// TIA Portal project "Impacchettatore" (V18)

(* hardware
DEVICE "S71500/ET200MP station_1"  S7-1500 station
   slot 0: "Telaio di montaggio_0"  Rack  6ES7 590-1***0-0AA0
   slot 1: "PLC_1"  CPU 1516-3 PN/DP  6ES7 516-3AN01-0AB0  V2.5
      slot 3: "Display CPU_1"  6ES7591-1BA00-0AA0
   slot 2: "DI 32x24VDC HF_1"  DI 32x24VDC HF  6ES7 521-1BL00-0AB0  V2.1
   slot 3: "DQ 32x24VDC/0.5A HF_1"  DQ 32x24VDC/0.5A HF  6ES7 522-1BL01-0AB0  V1.0
   slot 4: "AI 8xU/I/RTD/TC ST_1"  AI 8xU/I/RTD/TC ST  6ES7 531-7KF00-0AB0  V2.1
   slot 5: "AQ 4xU/I ST_1"  AQ 4xU/I ST  6ES7 532-5HD00-0AB0  V2.1
*)

// ===== PLC "PLC_1"  CPU 1516-3 PN/DP =====

VAR_GLOBAL   // PLC tag table "Tabella delle variabili standard"
   "slittaCentraleSu" AT %Q0.0 : Bool;
   "slittaCentraleGiu" AT %Q0.1 : Bool;
   "slittaSuperioreAvanti" AT %Q0.2 : Bool;
   "slittaSuperioreIndietro" AT %Q0.3 : Bool;
   "slittaEsternaSu" AT %Q0.4 : Bool;
   "motAvanti" AT %Q0.5 : Bool;
   "hg1" AT %Q0.6 : Bool;
   "hr2" AT %Q0.7 : Bool;
   "sensoreFondo" AT %I0.0 : Bool;
   "sensoreSopra" AT %I0.1 : Bool;
   "marcia" AT %I0.2 : Bool;
   "stop" AT %I0.3 : Bool;
   "inizializzazione" AT %I0.4 : Bool;
   "emergenza" AT %I0.5 : Bool;
   "readSlittaCentraleBasso" AT %I0.6 : Bool;
   "readSlittaCentraleAlto" AT %I0.7 : Bool;
   "readSlittaSuperioreIndietro" AT %I1.0 : Bool;
   "readSlittaSuperioreAvanti" AT %I1.1 : Bool;
   "readSlittaEsternaBasso" AT %I1.2 : Bool;
   "readSlittaEsternaAlto" AT %I1.3 : Bool;
END_VAR

DATA_BLOCK "DB_Comandi"   // DB1
{ S7_Optimized_Access := 'FALSE' }
VERSION : 0.1
   VAR
      btnInizializza : Bool;
      btnResetPezzi : Bool;
      btnStopNastro : Bool;
      btnSlittaLatGiu : Bool;
      btnSlittaLatSu : Bool;
      btnPistoneIndietro : Bool;
      btnPistoneAvanti : Bool;
      btnSlittaCentroGiu : Bool;
      btnSlittaCentroSu : Bool;
      btnNastro : Bool;
      bStop : Bool;
      bAuto : Bool;
      bMan : Bool;
      bReset : Bool;
      bEmergenza : Bool;
   END_VAR
BEGIN
END_DATA_BLOCK

DATA_BLOCK "DB_Stati"   // DB2
{ S7_Optimized_Access := 'FALSE' }
VERSION : 0.1
   VAR
      sAuto : Bool;
      sStop : Bool;
      sMan : Bool;
      sHome : Bool;
      sAttesastop : Bool;
      sEmergenza : Bool;
      bIni1 : Bool;
      bIni2 : Bool;
      bRip1 : Bool;
      bRip2 : Bool;
   END_VAR
BEGIN
END_DATA_BLOCK

DATA_BLOCK "DB_Tappe"   // DB3
{ S7_Optimized_Access := 'FALSE' }
VERSION : 0.1
   VAR
      tappeGemma : Int;
      tappeM1 : Int;
      tappeM2 : Int;
   END_VAR
BEGIN
END_DATA_BLOCK

DATA_BLOCK "DB_Variabili"   // DB4
{ S7_Optimized_Access := 'FALSE' }
VERSION : 0.1
   VAR
      timerResetPulsantiSTART : Bool;
      timerResetPulsantiDONE : Bool;
      timerResetPulsantiOUTPUT : Time;
      timerResetPulsantiDURATA : Time;
      timerSTART_1 : Bool;
      timerDONE_1 : Bool;
      timerOUTPUT_1 : Time;
      timerDURATA_1 : Time;
      timerSTART_2 : Bool;
      timerDONE_2 : Bool;
      timerOUTPUT_2 : Time;
      timerDURATA_2 : Time;
      timerSTART_3 : Bool;
      timerDONE_3 : Bool;
      timerOUTPUT_3 : Time;
      timerDURATA_3 : Time;
      timerSTART_4 : Bool;
      timerDONE_4 : Bool;
      timerOUTPUT_4 : Time;
      timerDURATA_4 : Time;
      statoLED : Bool;
      oSlittaEsterna : Bool;
      oPistoneIndietro : Bool;
      oPistoneAvanti : Bool;
      nCicli : Int;
      nPezzi : Int;
      oNastro : Bool;
      oSlittaSu : Bool;
      oLedVerde : Bool;
      oLedRosso : Bool;
      oSlittaGiu : Bool;
   END_VAR
BEGIN
END_DATA_BLOCK

// folder: System blocks/Program resources

DATA_BLOCK "timerResetPulsanti"   // DB5
{ S7_Optimized_Access := 'TRUE' }
AUTHOR : Simatic
FAMILY : IEC
NAME : IEC_TMR
VERSION : 1.0
// stored: InstanceOfName IEC_TIMER
"IEC_TIMER"
BEGIN
END_DATA_BLOCK

DATA_BLOCK "timer_1"   // DB6
{ S7_Optimized_Access := 'TRUE' }
AUTHOR : Simatic
FAMILY : IEC
NAME : IEC_TMR
VERSION : 1.0
// stored: InstanceOfName IEC_TIMER
"IEC_TIMER"
BEGIN
END_DATA_BLOCK

DATA_BLOCK "timer_2"   // DB7
{ S7_Optimized_Access := 'TRUE' }
AUTHOR : Simatic
FAMILY : IEC
NAME : IEC_TMR
VERSION : 1.0
// stored: InstanceOfName IEC_TIMER
"IEC_TIMER"
BEGIN
END_DATA_BLOCK

DATA_BLOCK "timer_3"   // DB8
{ S7_Optimized_Access := 'TRUE' }
AUTHOR : Simatic
FAMILY : IEC
NAME : IEC_TMR
VERSION : 1.0
// stored: InstanceOfName IEC_TIMER
"IEC_TIMER"
BEGIN
END_DATA_BLOCK

DATA_BLOCK "timer_4"   // DB9
{ S7_Optimized_Access := 'TRUE' }
AUTHOR : Simatic
FAMILY : IEC
NAME : IEC_TMR
VERSION : 1.0
// stored: InstanceOfName IEC_TIMER
"IEC_TIMER"
BEGIN
END_DATA_BLOCK

// folder: (top level)

FUNCTION "FC_Gemma" : Void   // FC1, SCL
{ S7_Optimized_Access := 'TRUE' }
VERSION : 0.1
BEGIN
   CASE "DB_Tappe".tappeGemma OF
       0:  // Stato di stop
           "DB_Stati".sStop := TRUE;
           IF "DB_Comandi".bAuto = TRUE THEN
               "DB_Tappe".tappeGemma := 1; //home
               "DB_Stati".sAttesastop := FALSE;
               "DB_Stati".sAuto := FALSE;
               "DB_Stati".sHome := TRUE;
               "DB_Stati".sMan := FALSE;
               "DB_Stati".sStop := FALSE;
           ELSE
               IF "DB_Comandi".bMan = TRUE THEN
                   "DB_Tappe".tappeGemma := 4; //manuale
                   "DB_Stati".sAttesastop := FALSE;
                   "DB_Stati".sAuto := FALSE;
                   "DB_Stati".sHome := FALSE;
                   "DB_Stati".sMan := TRUE;
                   "DB_Stati".sStop := FALSE;
               END_IF;
           END_IF;
       1:  // Stato di home
           IF "DB_Stati".bIni1 = TRUE AND "DB_Stati".bIni2 = TRUE THEN
               "DB_Tappe".tappeGemma := 2; //automatico
               "DB_Stati".sAttesastop := FALSE;
               "DB_Stati".sAuto := TRUE;
               "DB_Stati".sHome := FALSE;
               "DB_Stati".sMan := FALSE;
               "DB_Stati".sStop := FALSE;
           END_IF;
       2:  // Stato di automatico
           IF "DB_Comandi".bStop = TRUE THEN
               "DB_Tappe".tappeGemma := 3; //attesa stop
               "DB_Stati".sAttesastop := TRUE;
               "DB_Stati".sAuto := FALSE;
               "DB_Stati".sHome := FALSE;
               "DB_Stati".sMan := FALSE;
               "DB_Stati".sStop := FALSE;
           END_IF;
       3:  // Stato di attesaStop
           IF "DB_Stati".bRip1 = TRUE AND "DB_Stati".bRip2 = TRUE THEN
               "DB_Tappe".tappeGemma := 0; //stop
               "DB_Stati".sAttesastop := FALSE;
               "DB_Stati".sAuto := FALSE;
               "DB_Stati".sHome := FALSE;
               "DB_Stati".sMan := FALSE;
               "DB_Stati".sStop := TRUE;
           END_IF;
       4:  // Stato di manuale
           IF "DB_Comandi".bStop = TRUE THEN
               "DB_Tappe".tappeGemma := 0; //stop
               "DB_Stati".sAttesastop := FALSE;
               "DB_Stati".sAuto := FALSE;
               "DB_Stati".sHome := FALSE;
               "DB_Stati".sMan := FALSE;
               "DB_Stati".sStop := TRUE;
           END_IF;
       5:  // Stato di emergenza
           IF "DB_Comandi".bEmergenza = TRUE AND "DB_Stati".sEmergenza = TRUE THEN
               "DB_Tappe".tappeGemma := 0; //stop
               "DB_Stati".sEmergenza := FALSE;
               "DB_Stati".sAttesastop := FALSE;
               "DB_Stati".sAuto := FALSE;
               "DB_Stati".sHome := FALSE;
               "DB_Stati".sMan := FALSE;
               "DB_Stati".sStop := TRUE;
           END_IF;
   END_CASE;

   //gestione emergenza
   IF "DB_Comandi".bEmergenza = FALSE OR "emergenza" = FALSE THEN
       "DB_Tappe".tappeGemma := 5; //emergenza
       "DB_Stati".sEmergenza := TRUE;
       "DB_Stati".sAttesastop := FALSE;
       "DB_Stati".sAuto := FALSE;
       "DB_Stati".sHome := FALSE;
       "DB_Stati".sMan := FALSE;
       "DB_Stati".sStop := FALSE;
   END_IF;
END_FUNCTION

FUNCTION "FC_Grafcet" : Void   // FC2, SCL
{ S7_Optimized_Access := 'TRUE' }
VERSION : 0.1
BEGIN
   // Gestisco i comandi possibili in manuale o automatico

   "DB_Comandi".bAuto := "marcia";
   "DB_Comandi".bStop := "stop";
   "DB_Comandi".btnInizializza := "inizializzazione";

   IF "DB_Comandi".btnResetPezzi THEN
       "DB_Variabili".nCicli := 0;
       "DB_Variabili".nPezzi := 0;
       "DB_Comandi".btnResetPezzi := FALSE;
   END_IF;

   IF "sensoreFondo" = TRUE THEN
       "DB_Variabili".oLedRosso := TRUE;
   ELSE
       "DB_Variabili".oLedRosso := FALSE;
   END_IF;

   IF "DB_Stati".sEmergenza = TRUE THEN
       "DB_Variabili".oLedRosso := TRUE;
       "DB_Variabili".oLedVerde := TRUE;
   ELSE
       "DB_Variabili".oLedRosso := FALSE;
       "DB_Variabili".oLedVerde := FALSE;
   END_IF;

   IF "DB_Stati".sMan = TRUE THEN
       IF "DB_Comandi".btnNastro = TRUE AND "DB_Variabili".nPezzi < 3 AND "readSlittaCentraleBasso" = TRUE AND "sensoreFondo" = FALSE THEN
           "DB_Variabili".oNastro := TRUE;
           "DB_Comandi".btnNastro := FALSE;
           "DB_Variabili".timerSTART_1 := TRUE;
       END_IF;

       IF "DB_Comandi".btnStopNastro = TRUE AND "readSlittaCentraleBasso" = TRUE THEN
           "DB_Variabili".oNastro := FALSE;
           "DB_Comandi".btnStopNastro := FALSE;
       END_IF;

       IF "DB_Variabili".nPezzi = 3 AND "DB_Comandi".btnSlittaCentroSu = TRUE AND "sensoreFondo" = TRUE THEN
           "DB_Variabili".oSlittaGiu := FALSE;
           "DB_Variabili".oSlittaSu := TRUE;
           "DB_Comandi".btnSlittaCentroSu := FALSE;
           "DB_Variabili".nPezzi := 0;
           "DB_Variabili".nCicli += 1;
       END_IF;

       IF "DB_Comandi".btnSlittaCentroGiu = TRUE AND "DB_Variabili".nCicli <> 3 AND "sensoreSopra" = FALSE THEN
           "DB_Variabili".oSlittaSu := FALSE;
           "DB_Variabili".oSlittaGiu := TRUE;
           "DB_Comandi".btnSlittaCentroGiu := FALSE;
       END_IF;

       IF "DB_Comandi".btnPistoneAvanti = TRUE AND "DB_Variabili".nCicli = 3 AND "DB_Variabili".oSlittaEsterna = TRUE AND "readSlittaCentraleAlto" = TRUE AND "readSlittaEsternaAlto" = TRUE AND "sensoreSopra" = TRUE THEN
           "DB_Variabili".oPistoneIndietro := FALSE;
           "DB_Variabili".oPistoneAvanti := TRUE;
           "DB_Variabili".nCicli := 0;
           "DB_Comandi".btnPistoneAvanti := FALSE;
       END_IF;

       IF "DB_Comandi".btnPistoneIndietro = TRUE THEN
           "DB_Variabili".oPistoneAvanti := FALSE;
           "DB_Variabili".oPistoneIndietro := TRUE;
           "DB_Comandi".btnPistoneIndietro := FALSE;
       END_IF;

       IF "DB_Comandi".btnSlittaLatSu = TRUE THEN
           "DB_Variabili".oSlittaEsterna := TRUE;
           "DB_Comandi".btnSlittaLatSu := FALSE;
       END_IF;

       IF "DB_Comandi".btnSlittaLatGiu = TRUE THEN
           "DB_Variabili".oSlittaEsterna := FALSE;
           "DB_Comandi".btnSlittaLatGiu := FALSE;
       END_IF;

   END_IF;

   // Automatico solo iniziato
   // ELSIF "DB_Stati".sHome = TRUE THEN
   //     CASE "DB_Tappe".tappeM1 OF
   //         0:
   //             "DB_Stati".sAuto := TRUE;
   //             "DB_Variabili".oNastro := TRUE;
   //             "DB_Comandi".btnNastro := FALSE;
   //             "DB_Variabili".timerSTART_1 := TRUE;
   //     END_CASE;
   // END_IF;

   // Disabilito tutti i tasti in maniera tale che il bit non rimanga a TRUE
   "DB_Comandi".btnNastro := FALSE;
   "DB_Comandi".btnSlittaCentroGiu := FALSE;
   "DB_Comandi".btnSlittaCentroSu := FALSE;
   "DB_Comandi".btnPistoneIndietro := FALSE;
   "DB_Comandi".btnPistoneAvanti := FALSE;
   "DB_Comandi".btnSlittaLatGiu := FALSE;
   "DB_Comandi".btnSlittaLatSu := FALSE;


   IF "DB_Variabili".timerDONE_1 = TRUE THEN
       "DB_Variabili".timerDONE_1 := FALSE;
       "DB_Variabili".timerSTART_1 := FALSE;
       "DB_Variabili".oNastro := FALSE;
       "DB_Variabili".nPezzi += 3;
       "DB_Tappe".tappeM1 := 1;
   END_IF;
END_FUNCTION

FUNCTION "FC_ResetPulsanti" : Void   // FC3, SCL
{ S7_Optimized_Access := 'TRUE' }
VERSION : 0.1
BEGIN
   //simulo la pressione di un pulsante
   //fisico. dopo 500ms viene riportato a false
   //
   IF "DB_Comandi".bAuto = TRUE OR
       "DB_Comandi".bMan = TRUE OR
       "DB_Comandi".bReset = TRUE OR
       "DB_Comandi".bStop = TRUE THEN
       //faccio partire il timer
       "DB_Variabili".timerResetPulsantiSTART := TRUE;
   END_IF;
   //quando sono passati 500ms resetto i pulsanti
   IF "DB_Variabili".timerResetPulsantiDONE = TRUE THEN
       "DB_Comandi".bAuto := FALSE;
       "DB_Comandi".bMan := FALSE;
       "DB_Comandi".bReset := FALSE;
       "DB_Comandi".bStop := FALSE;
       //
       "DB_Variabili".timerResetPulsantiSTART := FALSE;
       "DB_Variabili".timerResetPulsantiDONE := FALSE;
   END_IF;
END_FUNCTION

FUNCTION "FC_Timer" : Void   // FC4, SCL
{ S7_Optimized_Access := 'TRUE' }
VERSION : 0.1
BEGIN
   "DB_Variabili".timerResetPulsantiDURATA := T#500ms;
   "timerResetPulsanti".TON(IN:="DB_Variabili".timerResetPulsantiSTART,
                            PT:="DB_Variabili".timerResetPulsantiDURATA,
                            Q=>"DB_Variabili".timerResetPulsantiDONE,
                            ET=>"DB_Variabili".timerResetPulsantiOUTPUT);
   //
   "DB_Variabili".timerDURATA_1 := T#7000ms;
   "timer_1".TON(IN:="DB_Variabili".timerSTART_1,
                 PT:="DB_Variabili".timerDURATA_1,
                 Q=>"DB_Variabili".timerDONE_1,
                 ET=>"DB_Variabili".timerOUTPUT_1);
   //
   "DB_Variabili".timerDURATA_2 := T#500ms;
   "timer_2".TON(IN:="DB_Variabili".timerSTART_2,
                 PT:="DB_Variabili".timerDURATA_2,
                 Q=>"DB_Variabili".timerDONE_2,
                 ET=>"DB_Variabili".timerOUTPUT_2);
   //
   "DB_Variabili".timerDURATA_3 := T#1500ms;
   "timer_3".TON(IN:="DB_Variabili".timerSTART_3,
                 PT:="DB_Variabili".timerDURATA_3,
                 Q=>"DB_Variabili".timerDONE_3,
                 ET=>"DB_Variabili".timerOUTPUT_3);
   //
   "DB_Variabili".timerDURATA_4 := T#200ms;
   "timer_4".TON(IN:="DB_Variabili".timerSTART_4,
                 PT:="DB_Variabili".timerDURATA_4,
                 Q=>"DB_Variabili".timerDONE_4,
                 ET=>"DB_Variabili".timerOUTPUT_4);
END_FUNCTION

FUNCTION "FC_Uscite" : Void   // FC5, SCL
{ S7_Optimized_Access := 'TRUE' }
VERSION : 0.1
BEGIN
   "motAvanti" := "DB_Variabili".oNastro;
   "slittaCentraleSu" := "DB_Variabili".oSlittaSu;
   "slittaCentraleGiu" := "DB_Variabili".oSlittaGiu;
   "slittaSuperioreAvanti" := "DB_Variabili".oPistoneAvanti;
   "slittaSuperioreIndietro" := "DB_Variabili".oPistoneIndietro;
   "slittaEsternaSu" := "DB_Variabili".oSlittaEsterna;
   "hg1" := "DB_Variabili".oLedVerde;
   "hr2" := "DB_Variabili".oLedRosso;

   IF (("DB_Stati".sAuto = TRUE AND "DB_Variabili".oNastro =
       TRUE)
       OR ("DB_Stati".sMan = TRUE AND "DB_Variabili".oNastro =
       TRUE))
       AND "DB_Stati".sEmergenza = FALSE THEN
       "motAvanti" := TRUE;
   ELSE
       "motAvanti" := FALSE;
   END_IF;

   IF (("DB_Stati".sAuto = TRUE AND "DB_Variabili".oSlittaGiu =
       TRUE)
       OR ("DB_Stati".sMan = TRUE AND "DB_Variabili".oSlittaGiu =
       TRUE))
       AND "DB_Variabili".oSlittaSu = FALSE
       AND "DB_Stati".sEmergenza = FALSE THEN
       "slittaCentraleGiu" := TRUE;
   ELSE
       "slittaCentraleGiu" := FALSE;
   END_IF;

   IF (("DB_Stati".sAuto = TRUE AND "DB_Variabili".oSlittaSu =
       TRUE)
       OR ("DB_Stati".sMan = TRUE AND "DB_Variabili".oSlittaSu =
       TRUE))
       AND "DB_Variabili".oSlittaGiu = FALSE
       AND "DB_Stati".sEmergenza = FALSE THEN
       "slittaCentraleSu" := TRUE;
   ELSE
       "slittaCentraleSu" := FALSE;
   END_IF;

   IF (("DB_Stati".sAuto = TRUE AND "DB_Variabili".oPistoneAvanti =
       TRUE)
       OR ("DB_Stati".sMan = TRUE AND "DB_Variabili".oPistoneAvanti =
       TRUE))
       AND "DB_Variabili".oPistoneIndietro = FALSE
       AND "DB_Stati".sEmergenza = FALSE THEN
       "slittaSuperioreAvanti" := TRUE;
   ELSE
       "slittaSuperioreAvanti" := FALSE;
   END_IF;

   IF (("DB_Stati".sAuto = TRUE AND "DB_Variabili".oPistoneIndietro =
       TRUE)
       OR ("DB_Stati".sMan = TRUE AND "DB_Variabili".oPistoneIndietro =
       TRUE))
       AND "DB_Variabili".oPistoneAvanti = FALSE
       AND "DB_Stati".sEmergenza = FALSE THEN
       "slittaSuperioreIndietro" := TRUE;
   ELSE
       "slittaSuperioreIndietro" := FALSE;
   END_IF;

   IF (("DB_Stati".sAuto = TRUE AND "DB_Variabili".oSlittaEsterna =
       TRUE)
       OR ("DB_Stati".sMan = TRUE AND "DB_Variabili".oSlittaEsterna =
       TRUE))
       AND "DB_Stati".sEmergenza = FALSE THEN
       "slittaEsternaSu" := TRUE;
   ELSE
       "slittaEsternaSu" := FALSE;
   END_IF;
END_FUNCTION

ORGANIZATION_BLOCK "Main"   // OB1, LAD, ProgramCycle
TITLE = "Main Program Sweep (Cycle)"
{ S7_Optimized_Access := 'TRUE' }
VERSION : 0.1
   VAR_INPUT
      Initial_Call : Bool;   // Initial call of this OB
      Remanence : Bool;   // =True, if remanent data are available
   END_VAR
   VAR_TEMP   // added for the SCL form of the ladder/FBD networks
      _w1 : Bool;
      _w2 : Bool;
      _w3 : Bool;
      _w4 : Bool;
   END_VAR
BEGIN

REGION Network 1
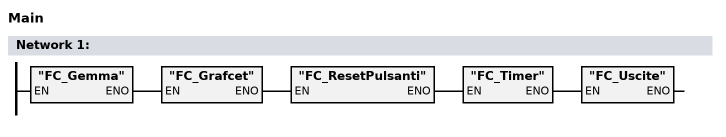
   RUNG wire#powerrail
      "FC_Gemma"()
      "FC_Grafcet"()
      "FC_ResetPulsanti"()
      "FC_Timer"()
      "FC_Uscite"()
   END_RUNG
   // the same network as SCL:
   "FC_Gemma"(ENO => #_w1);
   "FC_Grafcet"(EN := #_w1, ENO => #_w2);
   "FC_ResetPulsanti"(EN := #_w2, ENO => #_w3);
   "FC_Timer"(EN := #_w3, ENO => #_w4);
   IF #_w4 THEN "FC_Uscite"(); END_IF;
END_REGION
END_ORGANIZATION_BLOCK